(* IEC 61131-3 sources: sis-interlock-demo/pytests/golden/mini/src/POUs/Generated/F_SisIoKeys, 1 file *)

(* ---- F_SisIoKeys.decl.st ---- *)
// AUTO-GENERATED by cemgen 1.0.0 — не редактировать: правьте матрицу и запустите
//   python -m cemgen generate <файл матрицы .csv или .xlsx>
// Матрица: TEST-U301-CEM, объект U-301, ревизия 1 от 2026-10-16, SHA-256 сетки 9067fda96ae55e67
// Назначение: ключи и кнопка ПАЗ в образе ввода-вывода: пишет поля ключей разрешения байпасов и
//             обходов и кнопки «Сброс ПАЗ», если их теги заданы в матрице. TRUE — заданы все три
//             тега.
// Автор:      pytest; код — генератор cemgen
// Версия:     1.0.0
// Документ:   docs/DESIGN.md, раздел «10. Генератор cemgen»; docs/cause_effect_matrix.md
// ВНИМАНИЕ:   код демонстрационный и не предназначен для систем безопасности. Реальная ПАЗ требует
//             определения SIL, сертифицированных аппаратных и программных средств и валидации по
//             ГОСТ Р МЭК 61511.
FUNCTION F_SisIoKeys : BOOL
VAR_INPUT
    xBypassPermit   : BOOL;   // ключ «Разрешение байпасов»
    xOverridePermit : BOOL;   // ключ «Разрешение пусковых обходов»
    xResetPressed   : BOOL;   // кнопка «Сброс ПАЗ» нажата
END_VAR
VAR_IN_OUT
    stIo : ST_SisIo;          // образ ввода-вывода
END_VAR
